Staubli VAL3: HMI_prog.dtx

string sProgLsit
num nPageIndex
num nPageNum
string sSelProg
string sPageIndex
string sPageNum
public bool bBool[10]
bool bToSave
bool bBack
public bool bEditBool[9]
string sEditIndex
string sEditPage
string sSelTRAJ
num nEditPage
num nEditIndex
string sList[49]
bool bEditBack
bool bInsert
bool bCancel
string sSelType
string sSelItem
string sLastType
string sInsertList
num nType
public string sIF_Type[3]
public string sIF_Index[3]
num nIF_value[3]
num nProgType
string sInitialPassword = "55582930"
